Fanuc KAREL source: kt00871.KL

-- PROVISIONAL review KL for V1013-1; original PC SHA256 defd5aa28d5a4a5075d550951c1a032ecb8c7dad01c4eb3b2e123df1554fd0c5
-- Incomplete behavior may be omitted. Consult companion uncertainty JSON. Do not deploy.
PROGRAM KT00871
%NOLOCKGROUP
VAR
  R1 : REAL
  R2 : REAL
  OUT : REAL
BEGIN
  -- UNRESOLVED_PC offsets 5-16; opcodes 2E,23
  -- UNRESOLVED_PC offsets 21-32; opcodes 2E,23
  -- UNRESOLVED_PC offsets 37-48; opcodes 2E,23
  -- UNRESOLVED_PC offsets 53-64; opcodes 2E,23
  -- UNRESOLVED_PC offsets 69-85; opcodes 27,22,76,64,23
  -- UNRESOLVED_PC offsets 90-94; opcodes 7F
END KT00871
